Fanuc KAREL source: kb00040.KL

-- PROVISIONAL review KL for V770-1; original PC SHA256 d96ceee8a304480fd4b8db3f6e9089424216bf609741d1e0d04ef0412ade35da
-- Incomplete behavior may be omitted. Consult companion uncertainty JSON. Do not deploy.
PROGRAM KB00040
%NOLOCKGROUP
BEGIN
  -- UNRESOLVED_PC offsets 5-14; opcodes 3F,75
  -- UNRESOLVED_PC offsets 19-26; opcodes 9D,23
  -- UNRESOLVED_PC offsets 31-49; opcodes 27,22,2A,22,31
  -- UNRESOLVED_PC offsets 54-58; opcodes 7F
END KB00040
